TYPE "DT_ANA_CTRL_ALL"
VERSION : 0.1
   STRUCT
      MECH : "DT_ANA_CTRL_MECH";
   END_STRUCT;

END_TYPE

